FUNCTION_BLOCK SortingResetSequence (* The complete three step conveyor reset. *)
  (* Standard: 61499-2 *)
  (* Version 2.0, 2026-11-09, sorting2n, sorting2n *)
  PACKAGE Main;
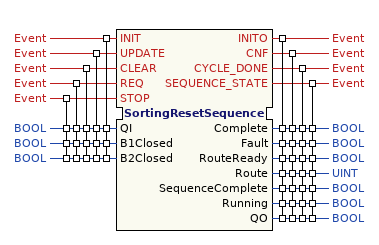
  EVENT_INPUT
    INIT WITH QI, B1Closed, B2Closed;
    UPDATE WITH QI, B1Closed, B2Closed;
    CLEAR WITH QI, B1Closed, B2Closed;
    REQ WITH QI, B1Closed, B2Closed;
    STOP WITH QI, B1Closed, B2Closed;
  END_EVENT
  EVENT_OUTPUT
    INITO WITH Complete, Fault, RouteReady, Route, SequenceComplete, Running, QO;
    CNF WITH Complete, Fault, RouteReady, Route, SequenceComplete, Running, QO;
    CYCLE_DONE WITH Complete, Fault, RouteReady, Route, SequenceComplete, Running, QO;
    SEQUENCE_STATE WITH Complete, Fault, RouteReady, Route, SequenceComplete, Running, QO;
  END_EVENT
  VAR_INPUT
    QI : BOOL := FALSE;
    B1Closed : BOOL;
    B2Closed : BOOL;
  END_VAR
  VAR_OUTPUT
    Complete : BOOL;
    Fault : BOOL;
    RouteReady : BOOL;
    Route : UINT := 0;
    SequenceComplete : BOOL;
    Running : BOOL := FALSE;
    QO : BOOL := FALSE;
  END_VAR
  FBS
    ResetSeq : SeqHead(PermStart := FALSE);
    TakeOwnership : SeqStep(TransStepId := 2);
    OwnershipTimeout : E_DELAY(DT := T#3s);
    CommandInitialPosition : SeqStep(Exceeded := TRUE, TransStepId := 3);
    Ready_CommandInitialPosition : E_SWITCH(G := TRUE);
    WaitInitialPosition : SeqStep(TransStepId := 4);
    InitialSettle : E_DELAY(DT := T#200ms);
    End : SeqTerminate;
    Frame : SortingCommandFrame;
    WriteCommands : SYMLINKMULTIVARSRC(QI := TRUE, NAME1 := '$${PATH:2}Conveyor.sc.lsp', NAME2 := '$${PATH:2}Branch1.sc.lsp', NAME3 := '$${PATH:2}Branch2.sc.lsp', NAME4 := '$${PATH:2}Stopper.sc.lsp'); {SET_ATTRIBUTE(Configuration.GenericFBType.InterfaceParams, Runtime.System#I:=4;VALUE${I$}:VTQINT,VTQINT,VTQINT,VTQINT)}
    Ownership : SortingOwnership;
    OwnerWrite : SYMLINKMULTIVARSRC(QI := TRUE, NAME1 := '$${PATH:2}Conveyor.sc.progLocalSel', NAME2 := '$${PATH:2}Branch1.sc.progLocalSel', NAME3 := '$${PATH:2}Branch2.sc.progLocalSel', NAME4 := '$${PATH:2}Stopper.sc.progLocalSel'); {SET_ATTRIBUTE(Configuration.GenericFBType.InterfaceParams, Runtime.System#I:=4;VALUE${I$}:VTQBOOL,VTQBOOL,VTQBOOL,VTQBOOL)}
    OwnerRead : SYMLINKMULTIVARDST(QI := TRUE, NAME1 := '$${PATH:2}Conveyor.sc.progLocal', NAME2 := '$${PATH:2}Branch1.sc.progLocal', NAME3 := '$${PATH:2}Branch2.sc.progLocal', NAME4 := '$${PATH:2}Stopper.sc.progLocal'); {SET_ATTRIBUTE(Configuration.GenericFBType.InterfaceParams, Runtime.System#I:=4;VALUE${I$}:VTQBOOL,VTQBOOL,VTQBOOL,VTQBOOL)}
    Home : SortingHomeConditions;
    HomeTimeout : E_DELAY(DT := T#2500ms);
  END_FBS
  EVENT_CONNECTIONS
    WaitInitialPosition.STEP_ENTER TO Home.C8FE616D2B744827;
    CommandInitialPosition.STEP_ENTER TO Ready_CommandInitialPosition.EI;
    OwnerRead.CNF TO Ownership.6D56496F53D1499B;
    Ownership.556ECCED2B7E4FE4 TO TakeOwnership.TRANS_REQ;
    Frame.91A08A19905E4AC8 TO WriteCommands.INIT;
    TakeOwnership.STEP_RESET TO OwnershipTimeout.STOP;
    Ownership.B3E6986DDAA841AB TO OwnerWrite.REQ;
    Ownership.4CD8C065E39641C9 TO OwnerWrite.INIT;
    ResetSeq.STATE_IND TO CNF;
    WaitInitialPosition.STEP_RESET TO HomeTimeout.STOP;
    OwnerRead.INITO TO Ownership.6D56496F53D1499B;
    InitialSettle.EO TO Home.858AFA5821D243F1;
    OwnershipTimeout.EO TO Home.BEAD4F12C24545AC;
    ResetSeq.STATE_IND TO SEQUENCE_STATE;
    Ready_CommandInitialPosition.EO1 TO CommandInitialPosition.TRANS_REQ;
    UPDATE TO ResetSeq.REQ_PERM;
    WaitInitialPosition.STEP_HOLD TO HomeTimeout.STOP;
    CLEAR TO Home.27094514BA434C7A;
    WriteCommands.INITO TO Ownership.D514169649844923;
    OwnerWrite.INITO TO OwnerRead.INIT;
    Home.C188F07096974982 TO ResetSeq.REQ_PERM;
    WaitInitialPosition.STEP_ENTER TO InitialSettle.START;
    WaitInitialPosition.STEP_RESET TO InitialSettle.STOP;
    WaitInitialPosition.STEP_HOLD TO InitialSettle.STOP;
    Frame.FEDD90899323480E TO WriteCommands.REQ;
    OwnerRead.INITO TO INITO;
    Home.199DF02180EA4007 TO CNF;
    STOP TO ResetSeq.RESET;
    HomeTimeout.EO TO Home.BEAD4F12C24545AC;
    WaitInitialPosition.STEP_LEAVE TO HomeTimeout.STOP;
    CommandInitialPosition.STEP_ENTER TO Frame.B00E6A8BE1EB4052;
    TakeOwnership.STEP_LEAVE TO OwnershipTimeout.STOP;
    TakeOwnership.STEP_ENTER TO OwnershipTimeout.START;
    UPDATE TO Home.F4871D28B0594017;
    OwnerRead.INITO TO Home.CE64267AAD124F8D;
    TakeOwnership.STEP_ENTER TO Ownership.8B11DD0F57C44878;
    Home.199DF02180EA4007 TO WaitInitialPosition.TRANS_REQ;
    WaitInitialPosition.STEP_LEAVE TO InitialSettle.STOP;
    INIT TO Frame.3E51AF3DA95F41C9;
    TakeOwnership.STEP_HOLD TO OwnershipTimeout.STOP;
    WaitInitialPosition.STEP_ENTER TO HomeTimeout.START;
    REQ TO ResetSeq.REQ_PERM;
    REQ TO ResetSeq.START;
  END_CONNECTIONS
  DATA_CONNECTIONS
    B2Closed TO Home.305FF7EA37BC4E0C;
    Frame.FD5B17DC6BEA4636 TO WriteCommands.VALUE3;
    Frame.E7BCFB58D0E944F4 TO WriteCommands.VALUE2;
    Ownership.AB3AFA1E5DB542BD TO OwnerWrite.VALUE3;
    Frame.1BE4F90CA0DE4A12 TO WriteCommands.VALUE1;
    OwnerRead.VALUE1 TO Ownership.3633AFB15F0E4D29;
    Ownership.AB3AFA1E5DB542BD TO OwnerWrite.VALUE4;
    Ownership.AB3AFA1E5DB542BD TO OwnerWrite.VALUE1;
    OwnerRead.VALUE4 TO Ownership.0CBD0A2278FC4256;
    B1Closed TO Home.6DF2726E50AE4D83;
    OwnerRead.VALUE2 TO Ownership.AFBF64D6B6724875;
    Home.74C9C2C856054ACB TO Fault;
    QI TO ResetSeq.PermStart;
    Ownership.3DD7BBA990934FB9 TO TakeOwnership.Exceeded;
    OwnerRead.VALUE3 TO Ownership.C6BAC61A3B114656;
    Frame.9F87DE883B874F73 TO WriteCommands.VALUE4;
    Home.097D9CE53785454A TO WaitInitialPosition.Exceeded;
    ResetSeq.SeqComplete TO SequenceComplete;
    ResetSeq.SeqComplete TO Complete;
    Ownership.AB3AFA1E5DB542BD TO OwnerWrite.VALUE2;
    ResetSeq.SeqRunning TO Running;
    QI TO QO;
  END_CONNECTIONS
  ADAPTER_CONNECTIONS
    ResetSeq.ISeqChain TO TakeOwnership.ISeqChainIn;
    WaitInitialPosition.ISeqChainOut TO End.ISeqChainIn;
    CommandInitialPosition.ISeqChainOut TO WaitInitialPosition.ISeqChainIn;
    TakeOwnership.ISeqChainOut TO CommandInitialPosition.ISeqChainIn;
  END_CONNECTIONS
END_FUNCTION_BLOCK
